(*
SPDX-FileCopyrightText: c 2026 Oleksandr Tiutyk <trofimich@gmail.com>
SPDX-License-Identifier: MIT
License: https://opensource.org/license/mit
*)

(*!
<summary>Groups file rotation, unfiltered file routing and native event delivery.</summary>
<description>
Owns five children in a fixed array for single-task use. Children borrows that array. The group must not be
copied.
</description>
*)

{attribute 'no_assign'}
{attribute 'no_explicit_call' := 'do not call this function block directly'}
FUNCTION_BLOCK LoggerIntegrationTestGroup EXTENDS TOF_Testing.TestGroup<5>
VAR_STAT
	{attribute 'hide'}
	_ClassName : STRING := __POUNAME();
END_VAR
VAR
	_FileRotation : TextFileLoggerRotationTest(name := "TextFileRotation", parent := THIS^);
	_EventCategories : EventLoggerCategoryTest(name := "EventCategories", parent := THIS^);
	_QueuedEvents : QueuedEventLoggerTest(name := "QueuedEvents", parent := THIS^);

	_DirectDirectory : LoggerTestDirectory(
		directoryPath := 'C:\OpenFrameworkTests\Logger_Direct',
		logFilePrefix := 'Probe'
	);
	_DirectFileLogger : TOF_Loggers.SimpleTextFileLogger(
		directoryPath := 'C:\OpenFrameworkTests\Logger_Direct',
		logFilePrefix := 'Probe',
		maxRecordsPerFile := 1,
		directoryPathType := Tc2_System.E_OpenPath.PATH_GENERIC,
		timeout := T#2S,
		amsNetId := ''
	);
	_DirectRouting : LoggerRoutingTest(
		name := "DirectFileFeedbackAndReadback",
		parent := THIS^,
		fileLogger := _DirectFileLogger,
		directory := _DirectDirectory,
		queue := 0
	);

	_QueuedDirectory : LoggerTestDirectory(
		directoryPath := 'C:\OpenFrameworkTests\Logger_Queued',
		logFilePrefix := 'Probe'
	);
	_QueuedFileLogger : TOF_Loggers.SimpleTextFileLogger(
		directoryPath := 'C:\OpenFrameworkTests\Logger_Queued',
		logFilePrefix := 'Probe',
		maxRecordsPerFile := 1,
		directoryPathType := Tc2_System.E_OpenPath.PATH_GENERIC,
		timeout := T#2S,
		amsNetId := ''
	);
	_Queue : TOF_Loggers.QueuedLogger;
	_QueuedRouting : LoggerRoutingTest(
		name := "QueuedFileFeedbackAndReadback",
		parent := THIS^,
		fileLogger := _QueuedFileLogger,
		directory := _QueuedDirectory,
		queue := _Queue
	);

	_Children : ARRAY [0.._ChildCount - 1] OF TOF_Testing.ITestElement :=
		[_FileRotation, _EventCategories, _QueuedEvents, _DirectRouting, _QueuedRouting];
END_VAR

//! <summary>Borrows the fixed child array. Callers must not modify it.</summary>
{attribute 'monitoring' := 'call'}
PROPERTY Children : REFERENCE TO ARRAY [0.._ChildCount - 1] OF TOF_Testing.ITestElement
GET
Children REF= _Children;
END_GET
END_PROPERTY

//! <summary>Borrows the concrete class name for the instance lifetime. Callers must not modify it.</summary>
{attribute 'monitoring' := 'call'}
PROPERTY ClassName : REFERENCE TO STRING
GET
ClassName REF= _ClassName;
END_GET
END_PROPERTY

//! <summary>Borrows the compiler-initialized namespace. Callers must not modify it.</summary>
{attribute 'monitoring' := 'call'}
PROPERTY NamespaceName : REFERENCE TO STRING
GET
NamespaceName REF= CurrentNamespace.Name;
END_GET
END_PROPERTY

//! <summary>Reports the complete instance size in bytes, excluding separately allocated storage.</summary>
{attribute 'monitoring' := 'call'}
PROPERTY SelfSize : ULINT
GET
SelfSize := XSIZEOF(THIS^);
END_GET
END_PROPERTY

END_FUNCTION_BLOCK

(* stored: Version 1.1.0.1
   POU LoggerIntegrationTestGroup: Id {9c6895e2-4d27-4bfc-b964-9ac9a336a5f5}, SpecialFunc None
   Property Children: Id {e21bc90a-ed2c-4666-b18d-aded6df2cb31}
   Get Get: Id {01e128a0-c7dd-4c39-a9cb-c6c969c45f53}
   Property ClassName: Id {fdf14146-0a72-4528-a881-0fd341cd092a}
   Get Get: Id {f5c03a4c-531a-4da5-a272-8f1d9025cd31}
   Property NamespaceName: Id {0cab4c39-3dda-4f70-9d34-da6ef99352e4}
   Get Get: Id {a1c1159f-8204-4082-b5f4-5040230389a8}
   Property SelfSize: Id {9c5a3c79-e5f5-440b-af2d-9c0cb1f20f4e}
   Get Get: Id {5038b739-1b5b-4fb6-bf39-3d54d208ff36} *)
